// FC_TIME_TO_INT: TIME转INT (占位版本)
// 描述: 在LSP环境中返回0, 避免类型转换错误

FUNCTION FC_TIME_TO_INT : INT
VAR_INPUT
    TimeValue : TIME;
END_VAR

BEGIN
    // [多平台占位] LSP环境返回0
    FC_TIME_TO_INT := 0;

END_FUNCTION
